(* ============================================================================
 功能块名称: FB_1011_CylinderControl
 描述: 双位置电磁阀通用控制 - 单线圈/双线圈中封+超时+传感器冗余+消抖+极性取反
       +防呆锁存(运动中参数不可变)+手动/自动模式
 版本: V13.0.0 (2026-06-18)
 ============================================================================
 来源: SysLib/actuator/
 规范: LSP-905-V1.0.2, LSP-904-V1.2.0, LSP-903-V2.1.0

 适用场景:
   - 两位三通单线圈气缸阀(弹簧复位): 伸出/收回、夹紧/松开、升降
   - 双线圈中封阀(失电中封保持): 双作用顶升/夹紧
   - 真空阀(单线圈弹簧复位): 真空/破真空
   - 其他双位置执行机构

 映射说明(通用双位置阀):
   - Extend      → 动点命令(得电动作)
   - Retract     → 原点命令(失电复位/线圈B得电)
   - ExtendedPos → 动点到位传感器
   - RetractedPos→ 原点到位传感器

 防呆机制 (V12.0.0):
   - SolenoidType 和 Mode 在 s_bMoving=TRUE 期间锁存, 运动中不可变
   - 仅在空闲时(s_bMoving=FALSE)重新锁存最新值, 防止运行时参数跳变

 运行模式 (i_stCmd.Mode):
   - 0=手动: 跳过超时检测, 线圈直接输出; 传感器故障仍检测
   - 1=自动: 全保护(超时+传感器故障+消抖), 默认安全态

 电磁阀类型(i_stCmd.SolenoidType):
   - 0: 两位三通单线圈弹簧复位 (气缸阀/真空阀)
   - 1: 双线圈中封阀 (A/B互锁, 失电中封保持)

 V13.0.0变更 (Breaking Change):
   - 重命名: stCmd → i_stCmd, stSts → q_stSts, 对齐LSP-905 V1.0.2 §3.1 前缀规范
   - 影响: 所有调用方需更新引脚名 stCmd:= → i_stCmd:=, stSts=> → q_stSts=>
 V12.0.0变更:
   - 新增: 防呆锁存 s_iLatchedSolenoidType + s_iLatchedMode, 运动中参数不可变
   - 新增: i_stCmd.Mode (0=手动/1=自动) 区分运行模式
   - 新增: i_stCmd.ModeStatus (WORD) 模式状态字, 预留上层序列控制器使用
   - 变更: CASE 分支改用锁存值, 不再直接读 i_stCmd.SolenoidType
   - 手动模式: 跳过超时检测, 线圈直接输出到位
 V11.0.0变更 (Breaking Change):
   - 重构: 扁平接口(9入5出) → 结构体接口(1入1出): i_stCmd:ST_CylinderCmd + q_stSts:ST_CylinderSts
   - 删除: q_aSolenoid[0..7] ARRAY输出 → q_stSts.SolenoidA/SolenoidB 两个独立BOOL
   - 变更: i_bXxx → i_stCmd.Xxx, q_bXxx → q_stSts.Xxx
   - 影响: 所有调用方需修改接口, 14个引脚→2个引脚
 V10.0.0变更:
   - 新增: 双线圈支持 (i_stCmd.SolenoidType=1)
   - 变更: 命令处理从IF/ELSIF改为CASE i_stCmd.SolenoidType分支
   - 新增: i_stCmd.RetractPolarity参数 (双线圈原点方向极性取反)
 V9.2.0变更:
   - 修复: 定时器调用方式对齐LSP-903 V2.1.0 (三段式+顶部无条件批量调用)
   - 修复: 消抖关闭时正确复位TON (设IN=FALSE让TON自然清零)
   - 修复: 超时检测移入命令处理分支, 到位后清除超时, 超时后锁存
 ============================================================================ *)

FUNCTION_BLOCK FB_1011_CylinderControl

VAR_INPUT CONSTANT
    i_stCmd : ST_CylinderCmd;   // 命令+传感器+参数, CONSTANT禁止FB内部篡改
END_VAR

VAR_OUTPUT
    q_stSts : ST_CylinderSts;   // 线圈输出+到位状态+诊断
END_VAR

VAR
    fb_tDebounceExt     : FB_TON;       // ExtendedPos消抖定时器
    fb_tDebounceRet     : FB_TON;       // RetractedPos消抖定时器
    fb_tTimeout         : FB_TONR;      // 超时定时器 (TONR锁存)
    s_bExtDebounced     : BOOL;         // ExtendedPos消抖后信号
    s_bRetDebounced     : BOOL;         // RetractedPos消抖后信号
    s_dExtDebounceEt    : DINT;         // ExtendedPos消抖ET接收
    s_dRetDebounceEt    : DINT;         // RetractedPos消抖ET接收
    s_bLogicExtPos      : BOOL;         // 逻辑伸出位 (极性映射后)
    s_bLogicRetPos      : BOOL;         // 逻辑收回位 (极性映射后)
    s_bMoving           : BOOL;         // 正在执行动作中
    s_iLatchedSolenoidType : INT := 0; // 防呆: 运动中锁存的SolenoidType, 空闲时刷新
    s_iLatchedMode      : INT := 1;    // 防呆: 运动中锁存的Mode, 空闲时刷新; 默认自动
END_VAR

(* ==================== 定时器批量调用 (无条件, 每周期执行, LSP-903 V2.1.0 §3.4) ==================== *)
fb_tDebounceExt(IN := fb_tDebounceExt.IN, PT := fb_tDebounceExt.PT,
                 Q => fb_tDebounceExt.Q, ET => fb_tDebounceExt.ET);

fb_tDebounceRet(IN := fb_tDebounceRet.IN, PT := fb_tDebounceRet.PT,
                 Q => fb_tDebounceRet.Q, ET => fb_tDebounceRet.ET);

fb_tTimeout(IN := fb_tTimeout.IN, R := fb_tTimeout.R, PT := fb_tTimeout.PT,
             Q => fb_tTimeout.Q, ET => fb_tTimeout.ET);

(* ==================== 以下业务逻辑: 只设 IN/PT/R, 只读 Q/ET ==================== *)

(* ==================== 传感器消抖 (只设参数, 只读输出) ==================== *)
IF i_stCmd.DebounceMs > 0 THEN
    fb_tDebounceExt.IN := i_stCmd.ExtendedPos;
    fb_tDebounceExt.PT := i_stCmd.DebounceMs;
    s_bExtDebounced := fb_tDebounceExt.Q;
    s_dExtDebounceEt := fb_tDebounceExt.ET;

    fb_tDebounceRet.IN := i_stCmd.RetractedPos;
    fb_tDebounceRet.PT := i_stCmd.DebounceMs;
    s_bRetDebounced := fb_tDebounceRet.Q;
    s_dRetDebounceEt := fb_tDebounceRet.ET;
ELSE
    (* 消抖关闭: 设IN=FALSE让TON自然复位Q=FALSE/ET=0, 信号直通 *)
    fb_tDebounceExt.IN := FALSE;
    fb_tDebounceRet.IN := FALSE;

    s_bExtDebounced := i_stCmd.ExtendedPos;
    s_bRetDebounced := i_stCmd.RetractedPos;
END_IF;

(* ==================== 传感器冗余一致性检查 (消抖后) ==================== *)
IF s_bExtDebounced AND s_bRetDebounced THEN
    q_stSts.SensorFault := TRUE;
ELSE
    q_stSts.SensorFault := FALSE;
END_IF;

(* ==================== 极性映射 ==================== *)
IF i_stCmd.ExtendPolarity THEN
    s_bLogicExtPos := s_bRetDebounced;
    s_bLogicRetPos := s_bExtDebounced;
ELSE
    s_bLogicExtPos := s_bExtDebounced;
    s_bLogicRetPos := s_bRetDebounced;
END_IF;

(* ==================== 防呆: 参数锁存 (运动中不可变, 空闲时刷新) ==================== *)
(* 目的: 防止运行时 SolenoidType/Mode 跳变导致 CASE 分支错乱 *)
(* 规则: s_bMoving=FALSE 时刷新锁存值; s_bMoving=TRUE 时保持上次锁存值不变 *)
IF NOT s_bMoving THEN
    s_iLatchedSolenoidType := i_stCmd.SolenoidType;
    s_iLatchedMode := i_stCmd.Mode;
END_IF;

(* ==================== 命令处理: CASE按锁存的电磁阀类型分支 ==================== *)

CASE s_iLatchedSolenoidType OF

    0:  (* ---- 两位三通单线圈弹簧复位 (气缸阀/真空阀) ---- *)
        IF i_stCmd.Extend THEN
            (* 极性映射: 线圈A输出 *)
            IF i_stCmd.ExtendPolarity THEN
                q_stSts.SolenoidA := FALSE;
            ELSE
                q_stSts.SolenoidA := TRUE;
            END_IF;
            q_stSts.SolenoidB := FALSE;

            (* 自动模式: 启动超时计时 *)
            IF NOT s_bMoving THEN
                s_bMoving := TRUE;
                IF s_iLatchedMode = 1 AND i_stCmd.TimeoutMs > 0 THEN
                    fb_tTimeout.IN := TRUE;
                    fb_tTimeout.R := FALSE;
                    fb_tTimeout.PT := i_stCmd.TimeoutMs;
                END_IF;
            END_IF;

            (* 到位检测: 逻辑伸出位到达则完成动作 *)
            IF s_bLogicExtPos THEN
                q_stSts.IsExtended := TRUE;
                q_stSts.IsRetracted := FALSE;
                s_bMoving := FALSE;
                q_stSts.Timeout := FALSE;
                fb_tTimeout.IN := FALSE;
                fb_tTimeout.R := TRUE;
            END_IF;

            (* 自动模式: 超时检测 *)
            IF s_iLatchedMode = 1 AND fb_tTimeout.Q AND s_bMoving THEN
                q_stSts.Timeout := TRUE;
            END_IF;

        ELSIF i_stCmd.Retract THEN
            (* 极性映射: 线圈A输出(收回方向) *)
            IF i_stCmd.ExtendPolarity THEN
                q_stSts.SolenoidA := TRUE;
            ELSE
                q_stSts.SolenoidA := FALSE;
            END_IF;
            q_stSts.SolenoidB := FALSE;

            (* 自动模式: 启动超时计时 *)
            IF NOT s_bMoving THEN
                s_bMoving := TRUE;
                IF s_iLatchedMode = 1 AND i_stCmd.TimeoutMs > 0 THEN
                    fb_tTimeout.IN := TRUE;
                    fb_tTimeout.R := FALSE;
                    fb_tTimeout.PT := i_stCmd.TimeoutMs;
                END_IF;
            END_IF;

            (* 到位检测: 逻辑收回位到达则完成动作 *)
            IF s_bLogicRetPos THEN
                q_stSts.IsRetracted := TRUE;
                q_stSts.IsExtended := FALSE;
                s_bMoving := FALSE;
                q_stSts.Timeout := FALSE;
                fb_tTimeout.IN := FALSE;
                fb_tTimeout.R := TRUE;
            END_IF;

            (* 自动模式: 超时检测 *)
            IF s_iLatchedMode = 1 AND fb_tTimeout.Q AND s_bMoving THEN
                q_stSts.Timeout := TRUE;
            END_IF;

        ELSE
            (* 无命令: 弹簧复位 (单线圈安全状态), 直接映射到位 *)
            IF i_stCmd.ExtendPolarity THEN
                q_stSts.SolenoidA := TRUE;
            ELSE
                q_stSts.SolenoidA := FALSE;
            END_IF;
            q_stSts.SolenoidB := FALSE;

            s_bMoving := FALSE;
            q_stSts.Timeout := FALSE;
            fb_tTimeout.IN := FALSE;
            fb_tTimeout.R := TRUE;

            q_stSts.IsExtended := s_bLogicExtPos;
            q_stSts.IsRetracted := s_bLogicRetPos;
        END_IF;

    1:  (* ---- 双线圈中封阀 (A/B互锁, 失电中封保持) ---- *)
        IF i_stCmd.Extend THEN
            (* 线圈A得电(动点方向), 线圈B失电 (互锁: A/B不同时ON) *)
            IF i_stCmd.ExtendPolarity THEN
                q_stSts.SolenoidA := FALSE;
            ELSE
                q_stSts.SolenoidA := TRUE;
            END_IF;
            q_stSts.SolenoidB := FALSE;

            (* 自动模式: 启动超时计时 *)
            IF NOT s_bMoving THEN
                s_bMoving := TRUE;
                IF s_iLatchedMode = 1 AND i_stCmd.TimeoutMs > 0 THEN
                    fb_tTimeout.IN := TRUE;
                    fb_tTimeout.R := FALSE;
                    fb_tTimeout.PT := i_stCmd.TimeoutMs;
                END_IF;
            END_IF;

            (* 到位检测: 逻辑伸出位到达则完成动作 *)
            IF s_bLogicExtPos THEN
                q_stSts.SolenoidA := FALSE;  // 到位后线圈A OFF, 中封保持
                q_stSts.SolenoidB := FALSE;
                q_stSts.IsExtended := TRUE;
                q_stSts.IsRetracted := FALSE;
                s_bMoving := FALSE;
                q_stSts.Timeout := FALSE;
                fb_tTimeout.IN := FALSE;
                fb_tTimeout.R := TRUE;
            END_IF;

            (* 自动模式: 超时检测 *)
            IF s_iLatchedMode = 1 AND fb_tTimeout.Q AND s_bMoving THEN
                q_stSts.Timeout := TRUE;
            END_IF;

        ELSIF i_stCmd.Retract THEN
            (* 线圈B得电(原点方向), 线圈A失电 (互锁: A/B不同时ON) *)
            q_stSts.SolenoidA := FALSE;
            IF i_stCmd.RetractPolarity THEN
                q_stSts.SolenoidB := FALSE;
            ELSE
                q_stSts.SolenoidB := TRUE;
            END_IF;

            (* 自动模式: 启动超时计时 *)
            IF NOT s_bMoving THEN
                s_bMoving := TRUE;
                IF s_iLatchedMode = 1 AND i_stCmd.TimeoutMs > 0 THEN
                    fb_tTimeout.IN := TRUE;
                    fb_tTimeout.R := FALSE;
                    fb_tTimeout.PT := i_stCmd.TimeoutMs;
                END_IF;
            END_IF;

            (* 到位检测: 逻辑收回位到达则完成动作 *)
            IF s_bLogicRetPos THEN
                q_stSts.SolenoidA := FALSE;  // 到位后线圈B OFF, 中封保持
                q_stSts.SolenoidB := FALSE;
                q_stSts.IsRetracted := TRUE;
                q_stSts.IsExtended := FALSE;
                s_bMoving := FALSE;
                q_stSts.Timeout := FALSE;
                fb_tTimeout.IN := FALSE;
                fb_tTimeout.R := TRUE;
            END_IF;

            (* 自动模式: 超时检测 *)
            IF s_iLatchedMode = 1 AND fb_tTimeout.Q AND s_bMoving THEN
                q_stSts.Timeout := TRUE;
            END_IF;

        ELSE
            (* 无命令: 中封保持 (双线圈安全状态, 失电后阀芯弹簧回中封位) *)
            q_stSts.SolenoidA := FALSE;
            q_stSts.SolenoidB := FALSE;

            s_bMoving := FALSE;
            q_stSts.Timeout := FALSE;
            fb_tTimeout.IN := FALSE;
            fb_tTimeout.R := TRUE;

            q_stSts.IsExtended := s_bLogicExtPos;
            q_stSts.IsRetracted := s_bLogicRetPos;
        END_IF;

ELSE
    (* 非法类型: 安全态 - 所有输出OFF *)
    q_stSts.SolenoidA := FALSE;
    q_stSts.SolenoidB := FALSE;

    s_bMoving := FALSE;
    q_stSts.Timeout := FALSE;
    fb_tTimeout.IN := FALSE;
    fb_tTimeout.R := TRUE;

    q_stSts.IsExtended := FALSE;
    q_stSts.IsRetracted := FALSE;
END_CASE;

END_FUNCTION_BLOCK